// TIA Portal V20 export
// export: Created 2026-10-19T18:07:48.9442604Z, ExportSetting None, DisplayName Totally Integrated Automation Portal, DisplayVersion V20 Update 6, DisplayName TIA Portal Openness, DisplayVersion V20 Update 6, DisplayName TIA Portal Version Control Interface, DisplayVersion V20 Update 6, DisplayName SINAMICS Startdrive Advanced, DisplayVersion V20 SP1, DisplayName SINAMICS Startdrive G130, G150, S120, S150, SINAMICS MV, G220, S200, S210, DisplayVersion V20 SP1, DisplayName SINAMICS Startdrive G110M, G120, G120C, G120D, G120P, G115D, DisplayVersion V20 SP1, DisplayName STEP 7 Professional, DisplayVersion V20 Update 6, DisplayName STEP 7 Safety, DisplayVersion V20 Update 2, DisplayName WinCC Basic/Comfort/Advanced, DisplayVersion V20 Update 6, DisplayName WinCC Unified, DisplayVersion V20 Update 6
VAR_GLOBAL   // PLC tag table "IND_360_Alibi"
   "AlibiGross_Byte(0)" AT %MB200 : Byte;
   "AlibiGross_Byte(1)" AT %MB201 : Byte;
   "AlibiGross_Byte(2)" AT %MB202 : Byte;
   "AlibiGross_Byte(3)" AT %MB203 : Byte;
   "AlibiNet_Byte(0)" AT %MB204 : Byte;
   "AlibiNet_Byte(1)" AT %MB205 : Byte;
   "AlibiNet_Byte(2)" AT %MB206 : Byte;
   "AlibiNet_Byte(3)" AT %MB207 : Byte;
   "AlibiTare_Byte(0)" AT %MB208 : Byte;
   "AlibiTare_Byte(1)" AT %MB209 : Byte;
   "AlibiTare_Byte(2)" AT %MB210 : Byte;
   "AlibiTare_Byte(3)" AT %MB211 : Byte;
   AlibiGross_Real AT %MD212 : Real;
   AlibiNet_Real AT %MD216 : Real;
   AlibiTare_Real AT %MD220 : Real;
END_VAR
